TYPE "FRK_HostEvents"
VERSION : 0.1
   STRUCT
      "Ring" : Array[1..32] of "ST_HostEvent";
      "RingHead" : Int;
      "Count" : Int;
      "Capacity" : Int;
      "Wrapped" : Bool;
   END_STRUCT;
END_TYPE
